(* IEC 61131-3 sources: nautilus/siemens/writer/testdata/dt, 2 files *)

(* ---- Fast.st ---- *)
(* A faster task: ramps over its dt-tag, an LREAL. *)
PROGRAM Fast
VAR_EXTERNAL
  FastDt : LREAL;
  Ramp : LREAL;
END_VAR
Ramp := Ramp + 2.0 * FastDt;
END_PROGRAM

(* ---- Main.st ---- *)
(* The main task: integrates over its own dt-tag (a REAL), and reads the
   fast task's (an LREAL), which makes that one a shared tag. *)
PROGRAM Main
VAR_EXTERNAL
  MainDtS : REAL;
  Hours : REAL;
  FastDt : LREAL;
  Seen : LREAL;
END_VAR
Hours := Hours + MainDtS / 3600.0;
Seen := FastDt;
END_PROGRAM
